Staubli VAL3: aioItem.pjx

--- aioItem.pjx ---
Parameters version=s8.10.3Cs9_BS2093 stackSize=5000 millimeterUnit=true
Program file=start.pgx
Program file=stop.pgx
Data file=aioItem.dtx

--- aioItem.dtx ---
public string sComment
public aio aAio

--- start.pgx ---
program start()
begin
end

--- stop.pgx ---
program stop()
begin
end
